RoboDK station: UR20_handgesture.rdk

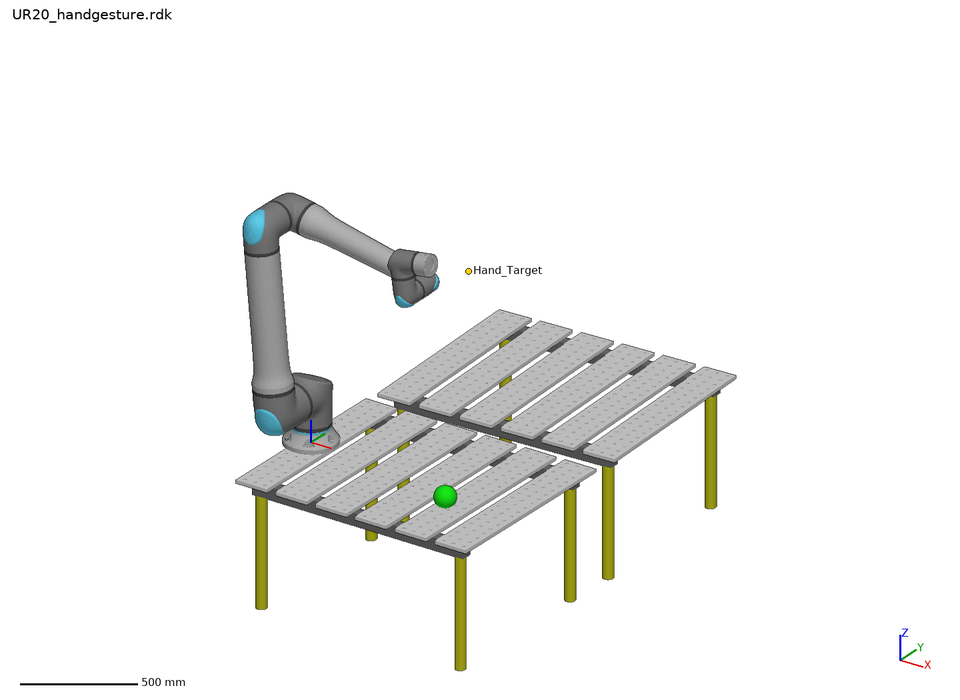
[picture v0: the station drawn from its stored meshes, robots at their saved joint values, targets as dots, program paths as lines]
Station hand_motion - Contactile (saved by RoboDK 6.0.6). Poses are relative to the parent item; angles as X-Y-Z fixed-axis rotations.
  - frame UR20 Base at (0, 0, 0) mm
    - robot UR20: 6 axes
        modified DH rows (alpha deg, a mm, theta deg, d mm): 0, 0, 0, 236.2; 90, 0, -180, 0; 0, 861.8, 0, 0; 0, 727.7, 0, 201.9; -90, 0, 0, 159.4; 90, 0, 180, 154.8
        joint limits [-360, -360, -360, -360, -360, -360] to [360, 360, 360, 360, 360, 360]; home [0, -90, -90, 0, 90, 0]; saved at [-0.125, -84.624, -106.704, 19.117, 90.125, 0]
    - target Hand_Target (Cartesian target) at (962.26, -203.23, 1157.29) mm, rotated rx -82.21 ry -0.02 rz -90 deg; joints [148.987, -31.705, 301.273, 90.432, 58.987, 180] of UR20
    - object Sphere D100mm at (829.04, -189.85, 50.02) mm, rotated rx -179.07 ry -0.46 rz 5.2 deg, size 100 x 100 x 100 mm, geometry from Sphere-D100mm.sld
  - object Table 1200x1000mm (Welding) at (543.39, 0, 0) mm, size 1193.8 x 965.2 x 609.6 mm, geometry from Table-1200x1000mm-Welding.sld
  - object Cube 50mm at (0, 0, 0) mm, size 100 x 100 x 100 mm, geometry from Cube-50mm.sld
  - object Table 1200x1000mm (Welding) at (534.06, 1058.97, 0) mm, rotated rx 0 ry 0 rz 2.59 deg, size 1193.8 x 965.2 x 609.6 mm, geometry from Table-1200x1000mm-Welding.sld
